// TIA Portal V20 export
Screen "MB150 first station LOADING STAND FIFO"  1276x673
  ScreenItem "线_1" at 0,65 size 1362x0  Type=HmiLine
  ScreenItem "permanentareaborderrectangle" at 0,0 size 0x0  Type=HmiRectangle
  ScreenItem "Button_Back" at 2,2 size 90x47  Type=HmiButton
  ScreenItem "OPMode4_Foreground_Blocked" at 1160,0 size 88x58  Type=HmiGraphicView
  ScreenItem "Title_OPOverview_ScreenOverview_X390_Y2" at 433,13 size 500x30  Type=HmiTextBox
  ScreenItem "Faceplate container_1" at 18,73 size 1239x577  Type=HmiFaceplateContainer
